(* IEC 61131-3 sources: plc-process-lib/src/POUs/Devices/FB_Valve, 28 files *)

(* ---- FB_Valve.decl.st ---- *)
// Назначение: запорная арматура двух видов. Задвижка с электроприводом (Motorized): выходы
//             «открывать» и «закрывать», стоп в промежутке, смена направления в ходе — через паузу
//             tReverse. Клапан с соленоидом (SolenoidEto, SolenoidEtc): одна катушка, пружинный
//             возврат. Открыть, закрыть, стоп от HMI и от автоматики; концевики ZSO/ZSC (или
//             положение по времени хода), контроль времени хода, «оба концевика», уход с концевика,
//             муфта ограничения момента, внешняя авария; Reset с окном tResetWindow; блокировки с
//             положением безопасности и первопричиной, разрешения по направлениям; режимы Auto,
//             Manual, Local, OutOfService; циклы и время работы привода в stRetain. Блокировка при одних
//             отказах контроля ведёт задвижку в положение безопасности (VLV-20); муфта открытия при
//             страгивании с седла — не заклинивание (VLV-21). Наследует FB_DeviceBase: тело — нормативный
//             порядок цикла (раздел 9.4 контракта).
// Автор:      kr0nsch
// Версия:     0.1.0
// Документ:   docs/fb/FB_Valve.md
FUNCTION_BLOCK FB_Valve EXTENDS FB_DeviceBase
VAR_INPUT
    xAutoOpen    : BOOL;             // запрос автоматики: TRUE — открыть, FALSE — закрыть
    xZso         : BOOL;             // концевик «открыто»
    xZsc         : BOOL;             // концевик «закрыто»
    xTorqueOpen  : BOOL;             // муфта (моментный выключатель) в сторону открытия
    xTorqueClose : BOOL;             // муфта в сторону закрытия
    xExtFault    : BOOL;             // авария привода: тепловое реле, обрыв фазы, авария интегрированного привода
    xLocal       : BOOL;             // «Местное» на приводе или шкафу
    xPowerOk     : BOOL := TRUE;     // напряжение питания привода
    wInterlock   : WORD := 16#0000;  // блокировки: бит = 1 — вести в eSafePos
    wPermitOpen  : WORD := 16#FFFF;  // разрешения на открытие: бит = 1 — разрешено
    wPermitClose : WORD := 16#FFFF;  // разрешения на закрытие: бит = 1 — разрешено
END_VAR
VAR_IN_OUT
    stCmd    : ST_ValveCmd;          // команды HMI/SCADA (GVL_Hmi.st<TAG>Cmd)
    stRetain : ST_DeviceRetain;      // режим, OOS, циклы, время работы привода (GVL_Persist.st<TAG>Retain)
END_VAR
VAR_IN_OUT CONSTANT
    stCfg : ST_ValveCfg;             // параметры (GVL_Persist.st<TAG>Cfg)
END_VAR
VAR_OUTPUT
    xQOpen  : BOOL;                  // Motorized: контактор «открывать»; соленоид — FALSE
    xQClose : BOOL;                  // Motorized: контактор «закрывать»; соленоид — FALSE
    xQCoil  : BOOL;                  // соленоид: катушка; Motorized — FALSE
    xOpened : BOOL;                  // положение «открыто» (по концевику или по времени хода)
    xClosed : BOOL;                  // положение «закрыто»
    stSts   : ST_ValveSts;           // состояние для HMI/SCADA
END_VAR
VAR
    stCfgLkg     : ST_ValveCfg;      // последняя корректная конфигурация (LKG, нормативно)
    // --- состояние и цель ---
    eState       : E_ValveState := E_ValveState.Unknown;        // состояние арматуры
    eTarget      : E_ValveState := E_ValveState.Intermediate;   // цель вызова: Open, Closed; Intermediate — «никуда»
    eManTarget   : E_ValveState := E_ValveState.Intermediate;   // цель Manual: последняя команда оператора
    eSolCmd      : E_ValveState := E_ValveState.Intermediate;  // соленоид: куда держит катушка; Intermediate — нет тока
    eLastEnd     : E_ValveState := E_ValveState.Unknown;        // последнее достигнутое крайнее положение (счёт циклов)
    eLastDir     : E_ValveState := E_ValveState.Intermediate;   // последнее включённое направление привода (выбег)
    xEndByLs     : BOOL;            // положение Open/Closed подтверждено своим концевиком (контроль ухода)
    // --- отказы: фиксируются до Reset (BothLimits — нет) ---
    xFltFailOpen  : BOOL;            // не открылась за tTravel
    xFltFailClose : BOOL;            // не закрылась за tTravel
    xFltPosLost   : BOOL;            // уход с концевика без команды
    xFltTorque    : BOOL;            // муфта в ходе
    xFltExt       : BOOL;            // внешняя авария
    xBothLimits   : BOOL;            // оба концевика дольше tLimitFilter (не фиксируется)
    xResetWin     : BOOL;            // идёт окно Reset: отказы снимаются, как только ушла причина
    // --- блокировки ---
    wIlkPrev      : WORD;            // блокировки после маски в прошлом вызове (первопричина)
    uiFirstOut    : UINT := GVL_Const.NO_FIRST_OUT;   // номер бита первой блокировки; NO_FIRST_OUT — нет
    // --- время работы привода ---
    xActPrev      : BOOL;            // в прошлом вызове был включён выход привода
    ltActAccum    : LTIME;           // накопитель времени работы привода: доля, меньшая 1 с
    // --- задержки (FB_Delay — единственный таймер библиотеки) ---
    fbTravel      : FB_Delay;        // время хода tTravel: от включения выхода (у соленоида — от смены цели)
    fbReverse     : FB_Delay;        // пауза перед реверсом tReverse
    fbRunOff      : FB_Delay;        // выбег привода: TRUE, пока выход включён, и ещё tReverse после снятия
    fbBoth        : FB_Delay;        // фильтр «оба концевика» tLimitFilter
    fbPosLost     : FB_Delay;        // фильтр ухода с концевика tLimitFilter
    fbResetWin    : FB_Delay;        // окно Reset tResetWindow
    // --- аварийный ход в положение безопасности при отказе контроля (VLV-20) ---
    xSafeMove     : BOOL;            // идёт аварийный ход по блокировке при отказе контроля (Motorized)
    xSafeMoveDone : BOOL;            // аварийный ход закончен: новый — после снятия блокировки или всех отказов
    eSafeDir      : E_ValveState := E_ValveState.Intermediate;   // направление аварийного хода: Opening, Closing
    fbSafeMove    : FB_Delay;        // время аварийного хода tTravel
    // --- страгивание с седла (VLV-21) ---
    xUnseatArmed  : BOOL;            // открытие началось с закрытого положения: муфта при страгивании не отказ
    fbUnseat      : FB_Delay;        // окно страгивания VLV_UNSEAT_BYPASS от начала открытия
    fbZscOff      : FB_Delay;        // ZSC замкнут или разомкнулся меньше tLimitFilter назад
    // --- сигналы и условия этого вызова: считает тело и шаги, читают следующие шаги ---
    xMotorized     : BOOL;           // электропривод (по LKG)
    xAtOpen        : BOOL;           // ZSO подключён и сработал
    xAtClose       : BOOL;           // ZSC подключён и сработал
    xTrqOpen       : BOOL;           // муфта открытия сработала (подключена, Motorized)
    xTrqClose      : BOOL;           // муфта закрытия сработала
    xRemote        : BOOL;           // режим Auto или Manual
    xSupervise     : BOOL;           // контроль концевиков: Auto/Manual и есть корректная Cfg
    xPosSup        : BOOL;           // контроль ухода с концевика: xSupervise и есть напряжение
    wIlk           : WORD;           // блокировки после маски
    xIlkAct        : BOOL;           // блокировка действует (Auto/Manual)
    wPermMissOpen  : WORD;           // недостающие разрешения на открытие
    wPermMissClose : WORD;           // недостающие разрешения на закрытие
    xMayOpen       : BOOL;           // открывать можно: разрешения есть или движение по блокировке
    xMayClose      : BOOL;           // закрывать можно
    xFaultAny      : BOOL;           // есть отказ (фиксированный или «оба концевика»)
    xDrive         : BOOL;           // ПЛК управляет выходами в этом вызове
    xEnterMove     : BOOL;           // в этом вызове началось движение (отсчёт tTravel заново)
END_VAR
VAR_TEMP
    eRes        : E_CmdResult;       // результат ProcessMode
    wPermMiss   : WORD;              // недостающие разрешения для текущего направления
    lrRemain_s  : LREAL;             // остаток времени хода, с
    udiRemain_s : UDINT;             // то же, целые секунды вверх
    xMaint      : BOOL;              // достигнут интервал ТО по циклам
    xAvailDev   : BOOL;              // готовность для автоматики (без учёта Cfg)
    wFltBits    : WORD;              // wFault
    wWrnBits    : WORD;              // wWarning
    wLowBits    : WORD;              // младший байт wStatus
    eDevSt      : E_Ne107Status;     // вклад устройства в NE 107
END_VAR

(* ---- CheckConfig.method.decl.st ---- *)
// Проверка конфигурации: биты wCfgErr арматуры (VLV_CFG_*). Только считает, ничего не меняет
METHOD PROTECTED CheckConfig : WORD
VAR_IN_OUT CONSTANT
    stCfgIn : ST_ValveCfg;   // проверяемая конфигурация
END_VAR
VAR
    wErr      : WORD;        // непройденные проверки
    xMotor    : BOOL;        // электропривод
    xSolenoid : BOOL;        // соленоид любого вида
END_VAR

(* ---- CheckConfig.method.impl.st ---- *)
xMotor := stCfgIn.eType = E_ValveType.Motorized;
xSolenoid := stCfgIn.eType = E_ValveType.SolenoidEto OR stCfgIn.eType = E_ValveType.SolenoidEtc;
IF NOT xMotor AND NOT xSolenoid THEN
    wErr := wErr OR GVL_Const.VLV_CFG_TYPE;
END_IF
IF stCfgIn.tTravel <= T#0S THEN
    wErr := wErr OR GVL_Const.VLV_CFG_TRAVEL;
END_IF
IF (stCfgIn.eSafePos <> E_ValveSafePos.Closed AND stCfgIn.eSafePos <> E_ValveSafePos.Open
    AND stCfgIn.eSafePos <> E_ValveSafePos.Stay)
   OR (xSolenoid AND stCfgIn.eSafePos = E_ValveSafePos.Stay)
THEN
    wErr := wErr OR GVL_Const.VLV_CFG_SAFE_POS;
END_IF
IF (stCfgIn.xCloseOnTorque AND NOT stCfgIn.xTorqueUsed) OR (xSolenoid AND stCfgIn.xTorqueUsed) THEN
    wErr := wErr OR GVL_Const.VLV_CFG_TORQUE;
END_IF
IF xMotor AND stCfgIn.tReverse <= T#0S THEN
    wErr := wErr OR GVL_Const.VLV_CFG_REVERSE;
END_IF
IF stCfgIn.tResetWindow <= T#0S THEN
    wErr := wErr OR GVL_Const.VLV_CFG_RESET;
END_IF
IF NOT CheckAlarmCfg(astCfg := stCfgIn.astAlarm) THEN
    wErr := wErr OR GVL_Const.VLV_CFG_ALARM;
END_IF
CheckConfig := wErr;

(* ---- CountOperations.method.decl.st ---- *)
// Шаг 6.9: циклы «открыто» и время работы привода в stRetain (параметр VAR_IN_OUT, R2).
// Шаг тела FB_Valve; внутренний: PROTECTED (правило L5 контракта), имя зарезервировано для наследников
METHOD PROTECTED CountOperations
VAR_IN_OUT
    stValveRet : ST_DeviceRetain;   // stRetain устройства
END_VAR

(* ---- CountOperations.method.impl.st ---- *)
// 6.9 Счётчики: цикл — вход в Open, если прошлое крайнее положение не Open; время работы — пока
//     включён выход привода (шаг не больше DT_ACCUM_MAX), целые секунды — в stRetain
IF eState = E_ValveState.Open AND eLastEnd <> E_ValveState.Open THEN
    stValveRet.udiOpCount := stValveRet.udiOpCount + 1;
    stValveRet.udiOpCountMaint := stValveRet.udiOpCountMaint + 1;
END_IF
IF eState = E_ValveState.Open OR eState = E_ValveState.Closed THEN
    eLastEnd := eState;
END_IF
IF xActPrev THEN
    ltActAccum := ltActAccum + MIN(ltDt, GVL_Const.DT_ACCUM_MAX);
END_IF
WHILE ltActAccum >= LTIME#1S DO
    ltActAccum := ltActAccum - LTIME#1S;
    stValveRet.udiOpTime_s := stValveRet.udiOpTime_s + 1;
    stValveRet.udiOpTimeMaint_s := stValveRet.udiOpTimeMaint_s + 1;
END_WHILE
xActPrev := xQOpen OR xQClose;

(* ---- CurrentTarget.method.impl.st ---- *)
IF eState = E_ValveState.Opening OR eState = E_ValveState.Open THEN
    CurrentTarget := E_ValveState.Open;
ELSIF eState = E_ValveState.Closing OR eState = E_ValveState.Closed THEN
    CurrentTarget := E_ValveState.Closed;
ELSIF eState = E_ValveState.Reversing THEN
    CurrentTarget := eTarget;
ELSE
    CurrentTarget := E_ValveState.Intermediate;
END_IF

(* ---- DriveToTarget.method.decl.st ---- *)
// Шаг 6.7: переходы движения к цели. Motorized: смена направления в ходе — через Reversing, стоп —
// Intermediate, встречное включение после остановки — не раньше tReverse (выбег); соленоид: смена цели —
// сразу другое направление; муфта в ходе — TorqueTrip, кроме страгивания с седла (VLV-21).
// Шаг тела FB_Valve; внутренний: PROTECTED (правило L5 контракта), имя зарезервировано для наследников
METHOD PROTECTED DriveToTarget
VAR
    xHoldOpen  : BOOL;   // открывать пока нельзя: «закрывать» снят меньше tReverse назад
    xHoldClose : BOOL;   // закрывать пока нельзя: «открывать» снят меньше tReverse назад
    xUnseating : BOOL;   // клин выходит из седла: муфта открытия — не заклинивание (VLV-21)
END_VAR

(* ---- DriveToTarget.method.impl.st ---- *)
// 6.7 Движение к цели. Motorized: смена направления в ходе — через Reversing; стоп — Intermediate.
//     Соленоид: смена цели в ходе — сразу другое направление, стопа нет
xMayOpen := xIlkAct OR wPermMissOpen = 0;
xMayClose := xIlkAct OR wPermMissClose = 0;
xEnterMove := FALSE;
//     выбег: встречное направление включается не раньше tReverse после снятия выхода — и после
//     остановки на концевике или по стопу, а не только при смене направления в ходе. Выходы здесь —
//     прошлого вызова; SetOutputs обновляет fbRunOff выходами этого вызова, поэтому отсчёт идёт ровно
//     от снятия выхода
fbRunOff(xIn := xQOpen OR xQClose, tOffDelay := stCfgLkg.tReverse, itfTime := itfTimeAct);
xHoldOpen := xMotorized AND fbRunOff.xOut AND eLastDir = E_ValveState.Closing;
xHoldClose := xMotorized AND fbRunOff.xOut AND eLastDir = E_ValveState.Opening;
//     страгивание с седла (VLV-21): усилие вырыва клина из седла больше усилия хода, муфта открытия срабатывает при
//     ещё замкнутом ZSC — это не заклинивание (в приводах — шунтирование моментного выключателя при страгивании).
//     Муфта открытия не контролируется, пока ZSC замкнут и ещё tLimitFilter после его размыкания (без ZSC — всё
//     окно), но не дольше VLV_UNSEAT_BYPASS от начала открытия с закрытого положения: клин, который не вышел из
//     седла, даёт TorqueTrip. Контроль заклинивания в ходе остаётся
IF eState <> E_ValveState.Opening THEN
    xUnseatArmed := FALSE;
END_IF
fbZscOff(xIn := xAtClose, tOffDelay := stCfgLkg.tLimitFilter, itfTime := itfTimeAct);
fbUnseat(xIn := xUnseatArmed AND eState = E_ValveState.Opening, tOnDelay := GVL_Const.VLV_UNSEAT_BYPASS,
         itfTime := itfTimeAct);
xUnseating := xUnseatArmed AND eState = E_ValveState.Opening AND NOT fbUnseat.xOut
              AND (fbZscOff.xOut OR NOT stCfgLkg.xZscUsed);
IF xDrive THEN
    IF eState = E_ValveState.Opening THEN
        IF xAtOpen THEN
            eState := E_ValveState.Open;
        ELSIF xTrqOpen AND NOT xUnseating THEN
            xFltTorque := TRUE;                // момент раньше концевика: заклинивание
            eState := E_ValveState.Fault;
        ELSIF eTarget = E_ValveState.Closed THEN
            IF xMotorized THEN
                eState := E_ValveState.Reversing;
            ELSIF xMayClose THEN
                eState := E_ValveState.Closing;
                xEnterMove := TRUE;
            END_IF
        ELSIF eTarget = E_ValveState.Intermediate AND xMotorized THEN
            eState := E_ValveState.Intermediate;
        END_IF
    ELSIF eState = E_ValveState.Closing THEN
        IF (xAtClose AND NOT stCfgLkg.xCloseOnTorque)
           OR (stCfgLkg.xCloseOnTorque AND xTrqClose AND (xAtClose OR NOT stCfgLkg.xZscUsed))
        THEN
            // по ZSC; при закрытии «по моменту» (клиновая задвижка) — только по муфте: ZSC стоит чуть
            // раньше посадки клина и выход не снимает, иначе задвижка не дожата. Муфта раньше
            // подключённого ZSC — не посадка, а заклинивание: TorqueTrip ниже
            eState := E_ValveState.Closed;
        ELSIF xTrqClose THEN
            xFltTorque := TRUE;
            eState := E_ValveState.Fault;
        ELSIF eTarget = E_ValveState.Open THEN
            IF xMotorized THEN
                eState := E_ValveState.Reversing;
            ELSIF xMayOpen THEN
                eState := E_ValveState.Opening;
                xEnterMove := TRUE;
            END_IF
        ELSIF eTarget = E_ValveState.Intermediate AND xMotorized THEN
            eState := E_ValveState.Intermediate;
        END_IF
    ELSIF eState = E_ValveState.Reversing THEN
        IF eTarget = E_ValveState.Intermediate THEN
            eState := E_ValveState.Intermediate;
        END_IF
    ELSIF eTarget = E_ValveState.Open AND eState <> E_ValveState.Open AND xMayOpen AND NOT xHoldOpen THEN
        // открытие с закрытого положения — окно страгивания от этого вызова
        xUnseatArmed := eState = E_ValveState.Closed;
        IF xUnseatArmed THEN
            fbUnseat.Preset(xValue := FALSE);
            fbUnseat(xIn := TRUE, tOnDelay := GVL_Const.VLV_UNSEAT_BYPASS, itfTime := itfTimeAct);
        END_IF
        eState := E_ValveState.Opening;
        xEnterMove := TRUE;
    ELSIF eTarget = E_ValveState.Closed AND eState <> E_ValveState.Closed AND xMayClose AND NOT xHoldClose THEN
        eState := E_ValveState.Closing;
        xEnterMove := TRUE;
    END_IF
END_IF

(* ---- FB_Valve.impl.st ---- *)
// 0. Первый вызов: число слотов тревог и тип устройства (до ProcessMode)
IF xFirstCall THEN
    uiAlarmCount := GVL_Const.VLV_ALARM_COUNT;
    eDevType := E_DeviceType.Valve;
END_IF

// 1. Время
BeginCycle();

// 2. Конфигурация (LKG)
IF AcceptCfg(wErr := CheckConfig(stCfgIn := stCfg)) THEN
    stCfgLkg := stCfg;
END_IF
// сигналы по LKG: концевик учитывается, только если подключён; муфта — только у Motorized
xMotorized := stCfgLkg.eType = E_ValveType.Motorized;
xAtOpen := stCfgLkg.xZsoUsed AND xZso;
xAtClose := stCfgLkg.xZscUsed AND xZsc;
xTrqOpen := xMotorized AND stCfgLkg.xTorqueUsed AND xTorqueOpen;
xTrqClose := xMotorized AND stCfgLkg.xTorqueUsed AND xTorqueClose;

// 3. Reset (метод ResetFaults; бит xReset сбрасывает RunAlarms в шаге 7)
ResetFaults(xRequest := xResetReq OR stCmd.stCommon.xReset);

// 4. Режим: вывод из работы — только когда арматура не движется
eRes := ProcessMode(xLocalSel := xLocal, xLocalSupported := TRUE,
                    xOosAllowed := eState <> E_ValveState.Opening AND eState <> E_ValveState.Closing
                                   AND eState <> E_ValveState.Reversing AND NOT xSafeMove,
                    stCmd := stCmd.stCommon, stRetain := stRetain);
IF eRes <> E_CmdResult.None THEN
    SetCmdResult(eResult := eRes);
END_IF

// 5. Условия вызова для шагов-методов; команды устройства (метод HandleCommands)
xRemote := eMode = E_DeviceMode.Auto OR eMode = E_DeviceMode.Manual;
wIlk := wInterlock AND stCfgLkg.wInterlockMask;
xIlkAct := xRemote AND wIlk <> 0;
wPermMissOpen := stCfgLkg.wPermitOpenMask AND NOT wPermitOpen;
wPermMissClose := stCfgLkg.wPermitCloseMask AND NOT wPermitClose;
xFaultAny := xFltFailOpen OR xFltFailClose OR xFltPosLost OR xFltTorque OR xFltExt OR xBothLimits;
HandleCommands(stValveCmd := stCmd, stValveRet := stRetain);

// 6. Логика по stCfgLkg: цель, контроль концевиков, состояние, движение, выходы, счётчики
SelectTarget();
SuperviseLimits();
TrackPosition();
DriveToTarget();
RunTravelTimers();
SafeMoveOnFault();
SetOutputs();
CountOperations(stValveRet := stRetain);

// 7. Тревоги (слоты E_ValveAlarm)
axAlmCond[E_ValveAlarm.FailToOpen] := xFltFailOpen;
axAlmCond[E_ValveAlarm.FailToClose] := xFltFailClose;
axAlmCond[E_ValveAlarm.BothLimits] := xBothLimits;
axAlmCond[E_ValveAlarm.PositionLost] := xFltPosLost;
axAlmCond[E_ValveAlarm.TorqueTrip] := xFltTorque;
axAlmCond[E_ValveAlarm.ExtFault] := xFltExt;
axAlmCond[E_ValveAlarm.InterlockAct] := xIlkAct;
RunAlarms(udiIdBase := stCfgLkg.udiAlarmIdBase, stCmd := stCmd.stCommon, astCfg := stCfgLkg.astAlarm);

// 8. Состояние
IF xRemote AND NOT xIlkAct AND eTarget = E_ValveState.Open AND eState <> E_ValveState.Open THEN
    wPermMiss := wPermMissOpen;
ELSIF xRemote AND NOT xIlkAct AND eTarget = E_ValveState.Closed AND eState <> E_ValveState.Closed THEN
    wPermMiss := wPermMissClose;
ELSE
    wPermMiss := 0;
END_IF
IF eState = E_ValveState.Opening OR eState = E_ValveState.Closing OR xSafeMove THEN
    // остаток до таймаута хода (аварийного хода), целые секунды вверх, не больше UINT_MAX
    IF xSafeMove THEN
        lrRemain_s := F_TimeToSec(tIn := fbSafeMove.tRemaining);
    ELSE
        lrRemain_s := F_TimeToSec(tIn := fbTravel.tRemaining);
    END_IF
    udiRemain_s := LREAL_TO_UDINT(lrRemain_s);
    IF UDINT_TO_LREAL(udiRemain_s) < lrRemain_s THEN
        udiRemain_s := udiRemain_s + 1;
    END_IF
    stSts.uiTravelRemain_s := UDINT_TO_UINT(MIN(udiRemain_s, UINT_TO_UDINT(GVL_Const.UINT_MAX)));
ELSE
    stSts.uiTravelRemain_s := 0;
END_IF
xMaint := stCfgLkg.udiMaintCycles > 0 AND stRetain.udiOpCountMaint >= stCfgLkg.udiMaintCycles;
wFltBits := SEL(xFltFailOpen, 0, GVL_Const.VLV_FLT_FAIL_TO_OPEN)
            OR SEL(xFltFailClose, 0, GVL_Const.VLV_FLT_FAIL_TO_CLOSE)
            OR SEL(xBothLimits, 0, GVL_Const.VLV_FLT_BOTH_LIMITS)
            OR SEL(xFltPosLost, 0, GVL_Const.VLV_FLT_POSITION_LOST)
            OR SEL(xFltTorque, 0, GVL_Const.VLV_FLT_TORQUE_TRIP)
            OR SEL(xFltExt, 0, GVL_Const.VLV_FLT_EXT_FAULT);
wWrnBits := SEL(xMaint, 0, GVL_Const.VLV_WRN_MAINT_CYCLES)
            OR SEL(xPowerOk, GVL_Const.VLV_WRN_POWER_LOST, 0)
            OR SEL(eMode = E_DeviceMode.Local AND wIlk <> 0, 0, GVL_Const.VLV_WRN_INTERLOCK_IN_LOCAL)
            OR SEL((eState = E_ValveState.Open AND NOT stCfgLkg.xZsoUsed)
                   OR (eState = E_ValveState.Closed AND NOT stCfgLkg.xZscUsed AND NOT stCfgLkg.xCloseOnTorque),
                   0, GVL_Const.VLV_WRN_POSITION_BY_TIME)
            OR SEL(eState = E_ValveState.Unknown, 0, GVL_Const.VLV_WRN_POSITION_UNKNOWN);
xAvailDev := eMode = E_DeviceMode.Auto AND wFltBits = 0 AND wIlk = 0 AND xPowerOk;
wLowBits := SEL(xOpened, 0, GVL_Const.VLV_STS_OPENED)
            OR SEL(xClosed, 0, GVL_Const.VLV_STS_CLOSED)
            OR SEL(eState = E_ValveState.Opening OR (xSafeMove AND eSafeDir = E_ValveState.Opening), 0,
                   GVL_Const.VLV_STS_OPENING)
            OR SEL(eState = E_ValveState.Closing OR (xSafeMove AND eSafeDir = E_ValveState.Closing), 0,
                   GVL_Const.VLV_STS_CLOSING)
            OR SEL(xIlkAct, 0, GVL_Const.VLV_STS_INTERLOCKED)
            OR SEL(wPermMiss <> 0, 0, GVL_Const.VLV_STS_PERMIT_MISSING)
            OR SEL(xTrqOpen OR xTrqClose, 0, GVL_Const.VLV_STS_TORQUE)
            OR SEL(xAvailDev AND xCfgEverOk, 0, GVL_Const.VLV_STS_AVAILABLE);
IF wFltBits <> 0 THEN
    eDevSt := E_Ne107Status.Failure;
ELSIF xMaint THEN
    eDevSt := E_Ne107Status.MaintenanceRequired;
ELSE
    eDevSt := E_Ne107Status.Good;
END_IF
stSts.eState := eState;
stSts.wInterlock := wIlk;
stSts.wPermitMissing := wPermMiss;
stSts.uiFirstOut := uiFirstOut;
stSts.wReserve := 0;
stSts.udiCycles := stRetain.udiOpCount;
stSts.udiCyclesMaint := stRetain.udiOpCountMaint;
stSts.rActTime_h := LREAL_TO_REAL(UDINT_TO_LREAL(stRetain.udiOpTime_s) / UDINT_TO_LREAL(GVL_Const.S_PER_H));
FinishCycle(eDevStatus := eDevSt, xAvailableDev := xAvailDev, wLow := wLowBits, wFaultBits := wFltBits,
            wWarnBits := wWrnBits, stCommon := stSts.stCommon);

(* ---- HandleCommands.method.decl.st ---- *)
// Шаг 5: команды HMI xClose > xOpen > xStop и xResetMaint; результат каждой — SetCmdResult. В Auto
// принятая команда переводит в Manual (оператор вмешался — автомат отпущен). Структуры — параметрами
// VAR_IN_OUT: метод не обращается к VAR_IN_OUT экземпляра (R2).
// Шаг тела FB_Valve; внутренний: PROTECTED (правило L5 контракта), имя зарезервировано для наследников
METHOD PROTECTED HandleCommands
VAR_IN_OUT
    stValveCmd : ST_ValveCmd;       // stCmd устройства: импульсы сбрасываются
    stValveRet : ST_DeviceRetain;   // stRetain устройства: режим, счётчики «с ТО»
END_VAR
VAR
    eCmdTgt : E_ValveState := E_ValveState.Intermediate;   // цель команды; Intermediate — стоп
    eResCmd : E_CmdResult := E_CmdResult.None;             // результат команды
END_VAR

(* ---- HandleCommands.method.impl.st ---- *)
IF stValveCmd.xClose OR stValveCmd.xOpen OR stValveCmd.xStop THEN
    IF stValveCmd.xClose THEN
        eCmdTgt := E_ValveState.Closed;
    ELSIF stValveCmd.xOpen THEN
        eCmdTgt := E_ValveState.Open;
    ELSE
        eCmdTgt := E_ValveState.Intermediate;
    END_IF
    IF NOT xRemote THEN
        eResCmd := E_CmdResult.RejectedMode;
    ELSIF eCmdTgt = E_ValveState.Intermediate THEN
        // стоп: только у электропривода; безопасен, поэтому без проверки Cfg и отказов
        IF NOT xMotorized THEN
            eResCmd := E_CmdResult.RejectedNotSupported;
        ELSIF xIlkAct THEN
            eResCmd := E_CmdResult.RejectedInterlock;
        ELSE
            eResCmd := E_CmdResult.Accepted;
        END_IF
    ELSIF NOT xCfgEverOk THEN
        eResCmd := E_CmdResult.RejectedCfg;
    ELSIF xFaultAny THEN
        eResCmd := E_CmdResult.RejectedFault;
    ELSIF xIlkAct THEN
        eResCmd := E_CmdResult.RejectedInterlock;
    ELSIF (eCmdTgt = E_ValveState.Open AND wPermMissOpen <> 0)
          OR (eCmdTgt = E_ValveState.Closed AND wPermMissClose <> 0)
    THEN
        eResCmd := E_CmdResult.RejectedPermit;
    ELSIF NOT xPowerOk THEN
        eResCmd := E_CmdResult.RejectedInhibit;
    ELSE
        eResCmd := E_CmdResult.Accepted;
    END_IF
    IF eResCmd = E_CmdResult.Accepted THEN
        // Auto -> Manual (хук: цель := текущее направление); в Manual режим не меняется
        SwitchRemoteMode(eNew := E_DeviceMode.Manual, stRetain := stValveRet);
        eManTarget := eCmdTgt;
    END_IF
    SetCmdResult(eResult := eResCmd);
END_IF
stValveCmd.xOpen := FALSE;
stValveCmd.xClose := FALSE;
stValveCmd.xStop := FALSE;
IF stValveCmd.xResetMaint THEN
    stValveRet.udiOpCountMaint := 0;
    stValveRet.udiOpTimeMaint_s := 0;
    SetCmdResult(eResult := E_CmdResult.Accepted);
    stValveCmd.xResetMaint := FALSE;
END_IF

(* ---- LimitPosition.method.decl.st ---- *)
// Положение по концевикам (с учётом «подключён»): только ZSO — Open, только ZSC — Closed, оба —
// Unknown; ни одного — Intermediate, а без концевиков — Unknown. Старт ПЛК и снятие отказа.
// Внутренний шаг устройства: PROTECTED (правило L5 контракта), имя зарезервировано для наследников
METHOD PROTECTED LimitPosition : E_ValveState
VAR
    xOpenLs  : BOOL;   // ZSO подключён и сработал
    xCloseLs : BOOL;   // ZSC подключён и сработал
END_VAR

(* ---- LimitPosition.method.impl.st ---- *)
xOpenLs := stCfgLkg.xZsoUsed AND xZso;
xCloseLs := stCfgLkg.xZscUsed AND xZsc;
IF xOpenLs AND xCloseLs THEN
    LimitPosition := E_ValveState.Unknown;
ELSIF xOpenLs THEN
    LimitPosition := E_ValveState.Open;
ELSIF xCloseLs THEN
    LimitPosition := E_ValveState.Closed;
ELSIF stCfgLkg.xZsoUsed OR stCfgLkg.xZscUsed THEN
    LimitPosition := E_ValveState.Intermediate;
ELSE
    LimitPosition := E_ValveState.Unknown;
END_IF

(* ---- OnModeChanged.method.decl.st ---- *)
// Хук смены режима: сначала база (SUPER^); переход в Manual — цель := текущее направление или
// положение (арматура не дёргается); вход в OutOfService снимает зафиксированные отказы и
// первопричину. VAR_IN_OUT устройства не трогает (R2)
METHOD PROTECTED OnModeChanged
VAR_INPUT
    eOld : E_DeviceMode;   // режим до смены
    eNew : E_DeviceMode;   // новый режим
END_VAR

(* ---- OnModeChanged.method.impl.st ---- *)
SUPER^.OnModeChanged(eOld := eOld, eNew := eNew);
IF eNew = E_DeviceMode.Manual THEN
    eManTarget := CurrentTarget();
END_IF
IF eNew = E_DeviceMode.OutOfService THEN
    xFltFailOpen := FALSE;
    xFltFailClose := FALSE;
    xFltPosLost := FALSE;
    xFltTorque := FALSE;
    xFltExt := FALSE;
    xResetWin := FALSE;
    uiFirstOut := GVL_Const.NO_FIRST_OUT;
END_IF

(* ---- ResetFaults.method.decl.st ---- *)
// Шаг 3: Reset. Результат Accepted сразу; в окне tResetWindow зафиксированные отказы снимаются, как
// только ушла их причина (ход и положение — сразу: привод стоит); если к концу окна отказ остался —
// второй результат RejectedFault. Первопричина блокировки снимается.
// Шаг тела FB_Valve; внутренний: PROTECTED (правило L5 контракта), имя зарезервировано для наследников
METHOD PROTECTED ResetFaults
VAR_INPUT
    xRequest : BOOL;   // Reset() или stCmd.stCommon.xReset в этом вызове
END_VAR

(* ---- ResetFaults.method.impl.st ---- *)
IF xRequest THEN
    uiFirstOut := GVL_Const.NO_FIRST_OUT;
    SetCmdResult(eResult := E_CmdResult.Accepted);
    IF xFltFailOpen OR xFltFailClose OR xFltPosLost OR xFltTorque OR xFltExt THEN
        xResetWin := TRUE;
        fbResetWin.Preset(xValue := FALSE);
    END_IF
END_IF
fbResetWin(xIn := xResetWin, tOnDelay := stCfgLkg.tResetWindow, itfTime := itfTimeAct);
IF xResetWin THEN
    // отказы хода и положения: привод стоит, причина в прошлом — снимаются сразу
    xFltFailOpen := FALSE;
    xFltFailClose := FALSE;
    xFltPosLost := FALSE;
    IF NOT xTrqOpen AND NOT xTrqClose THEN
        xFltTorque := FALSE;
    END_IF
    IF NOT xExtFault THEN
        xFltExt := FALSE;
    END_IF
    IF NOT xFltTorque AND NOT xFltExt THEN
        xResetWin := FALSE;
    ELSIF fbResetWin.xOut THEN
        SetCmdResult(eResult := E_CmdResult.RejectedFault);
        xResetWin := FALSE;
    END_IF
END_IF

(* ---- RunTravelTimers.method.impl.st ---- *)
//     пауза реверса: отсчёт с входа в Reversing, затем направление по цели
fbReverse(xIn := eState = E_ValveState.Reversing, tOnDelay := stCfgLkg.tReverse, itfTime := itfTimeAct);
IF eState = E_ValveState.Reversing AND fbReverse.xOut THEN
    IF eTarget = E_ValveState.Open AND xMayOpen THEN
        eState := E_ValveState.Opening;
        xEnterMove := TRUE;
    ELSIF eTarget = E_ValveState.Closed AND xMayClose THEN
        eState := E_ValveState.Closing;
        xEnterMove := TRUE;
    ELSE
        eState := E_ValveState.Intermediate;
    END_IF
END_IF
//     время хода: отсчёт заново с каждого начала движения. Концевик положения подключён (у
//     закрытия — или закрытие по моменту) — таймаут = отказ; не подключён — положение по времени
IF xEnterMove THEN
    fbTravel.Preset(xValue := FALSE);
END_IF
fbTravel(xIn := eState = E_ValveState.Opening OR eState = E_ValveState.Closing, tOnDelay := stCfgLkg.tTravel,
         itfTime := itfTimeAct);
IF fbTravel.xOut THEN
    IF eState = E_ValveState.Opening THEN
        IF stCfgLkg.xZsoUsed THEN
            xFltFailOpen := TRUE;
            eState := E_ValveState.Fault;
        ELSE
            eState := E_ValveState.Open;
        END_IF
    ELSIF eState = E_ValveState.Closing THEN
        IF stCfgLkg.xZscUsed OR stCfgLkg.xCloseOnTorque THEN
            xFltFailClose := TRUE;
            eState := E_ValveState.Fault;
        ELSE
            eState := E_ValveState.Closed;
        END_IF
    END_IF
END_IF

//     крайнее положение подтверждено концевиком (по времени хода и «по моменту» — нет): только
//     такое положение контролируется на уход с концевика
IF (eState = E_ValveState.Open AND xAtOpen) OR (eState = E_ValveState.Closed AND xAtClose) THEN
    xEndByLs := TRUE;
ELSIF eState <> E_ValveState.Open AND eState <> E_ValveState.Closed THEN
    xEndByLs := FALSE;
END_IF

(* ---- SafeMoveOnFault.method.decl.st ---- *)
// Шаг 6.7а (VLV-20): аварийный ход в положение безопасности по блокировке, когда отказали только средства
// контроля (BothLimits, PositionLost, FailToOpen, FailToClose), а привод исправен: защита важнее диагностики.
// Только Motorized (соленоид при отказе уходит на пружину, A-10), с положением безопасности Open или Closed; не
// при внешней аварии, муфте, без напряжения и без корректной Cfg. Концевикам при отказе контроля верить нельзя:
// ход заканчивается по согласованному концевику положения безопасности (свой замкнут, встречный нет), по муфте в
// этом направлении или через tTravel. Пока блокировка и отказ держатся, ход не повторяется. Начало — после выбега
// встречного направления (VLV-05).
// Шаг тела FB_Valve; внутренний: PROTECTED (правило L5 контракта), имя зарезервировано для наследников
METHOD PROTECTED SafeMoveOnFault
VAR
    xMayMove : BOOL;   // аварийный ход допустим в этом вызове
    xEnd     : BOOL;   // аварийный ход закончен в этом вызове
END_VAR

(* ---- SafeMoveOnFault.method.impl.st ---- *)
xMayMove := xMotorized AND xIlkAct AND xFaultAny AND xCfgEverOk AND xPowerOk AND NOT xFltExt AND NOT xFltTorque
            AND (stCfgLkg.eSafePos = E_ValveSafePos.Open OR stCfgLkg.eSafePos = E_ValveSafePos.Closed);
IF NOT xMayMove THEN
    xSafeMove := FALSE;
    IF NOT (xIlkAct AND xFaultAny) THEN
        // блокировка или отказы сняты: следующий эпизод — новый аварийный ход
        xSafeMoveDone := FALSE;
    END_IF
ELSIF NOT xSafeMove AND NOT xSafeMoveDone THEN
    IF stCfgLkg.eSafePos = E_ValveSafePos.Closed AND NOT (fbRunOff.xOut AND eLastDir = E_ValveState.Opening) THEN
        eSafeDir := E_ValveState.Closing;
        xSafeMove := TRUE;
    ELSIF stCfgLkg.eSafePos = E_ValveSafePos.Open AND NOT (fbRunOff.xOut AND eLastDir = E_ValveState.Closing) THEN
        eSafeDir := E_ValveState.Opening;
        xSafeMove := TRUE;
    END_IF
    IF xSafeMove THEN
        fbSafeMove.Preset(xValue := FALSE);
    END_IF
END_IF
fbSafeMove(xIn := xSafeMove, tOnDelay := stCfgLkg.tTravel, itfTime := itfTimeAct);
IF xSafeMove THEN
    IF eSafeDir = E_ValveState.Closing THEN
        xEnd := (xAtClose AND NOT xAtOpen) OR xTrqClose;
    ELSE
        xEnd := (xAtOpen AND NOT xAtClose) OR xTrqOpen;
    END_IF
    IF xEnd OR fbSafeMove.xOut THEN
        xSafeMove := FALSE;
        xSafeMoveDone := TRUE;
    END_IF
END_IF

(* ---- SelectTarget.method.decl.st ---- *)
// Шаг 6.1–6.2: цель вызова (Auto — запрос автоматики, Manual — команда оператора, Local/OOS — нет,
// блокировка — положение безопасности) и первопричина блокировки.
// Шаг тела FB_Valve; внутренний: PROTECTED (правило L5 контракта), имя зарезервировано для наследников
METHOD PROTECTED SelectTarget
VAR
    wBit  : WORD;   // бит при поиске первопричины
    uiBit : UINT;   // номер бита
END_VAR

(* ---- SelectTarget.method.impl.st ---- *)
// 6.1 Цель: Auto — по запросу автоматики, Manual — по команде оператора, Local/OOS — нет;
//     блокировка (Auto/Manual) — положение безопасности (Stay — стоп)
IF eMode = E_DeviceMode.Auto THEN
    IF xAutoOpen THEN
        eTarget := E_ValveState.Open;
    ELSE
        eTarget := E_ValveState.Closed;
    END_IF
ELSIF eMode = E_DeviceMode.Manual THEN
    eTarget := eManTarget;
ELSE
    eTarget := E_ValveState.Intermediate;
END_IF
IF xIlkAct THEN
    IF stCfgLkg.eSafePos = E_ValveSafePos.Open THEN
        eTarget := E_ValveState.Open;
    ELSIF stCfgLkg.eSafePos = E_ValveSafePos.Closed THEN
        eTarget := E_ValveState.Closed;
    ELSE
        eTarget := E_ValveState.Intermediate;
    END_IF
    // блокировка не фиксируется: после её снятия Manual остаётся в положении безопасности
    IF eMode = E_DeviceMode.Manual THEN
        eManTarget := eTarget;
    END_IF
END_IF

// 6.2 Первопричина: при переходе слова блокировок из 0 в не 0 — номер младшего взведённого бита
//     (держится до Reset или входа в OutOfService). Цикл конечен: wIlk <> 0
IF wIlkPrev = 0 AND wIlk <> 0 AND eMode <> E_DeviceMode.OutOfService THEN
    wBit := 1;
    uiBit := 0;
    WHILE (wIlk AND wBit) = 0 DO
        wBit := SHL(wBit, 1);
        uiBit := uiBit + 1;
    END_WHILE
    uiFirstOut := uiBit;
END_IF
wIlkPrev := wIlk;

(* ---- SetOutputs.method.decl.st ---- *)
// Шаг 6.8: выходы привода и катушки, положение для логики. Без управления и при отказе выходы сняты,
// катушка обесточена (положение пружины); при отказе контроля — аварийный ход по блокировке (VLV-20).
// Шаг тела FB_Valve; внутренний: PROTECTED (правило L5 контракта), имя зарезервировано для наследников
METHOD PROTECTED SetOutputs
VAR
    xOutEn : BOOL;   // выходы разрешены
END_VAR

(* ---- SetOutputs.method.impl.st ---- *)
// 6.8 Выходы. Без управления и при отказе выходы сняты, катушка обесточена (положение пружины)
IF NOT xDrive OR eState = E_ValveState.Fault OR xMotorized THEN
    eSolCmd := E_ValveState.Intermediate;
ELSIF eState = E_ValveState.Opening OR (eState = E_ValveState.Open AND eTarget = E_ValveState.Open) THEN
    eSolCmd := E_ValveState.Open;
ELSIF eState = E_ValveState.Closing OR (eState = E_ValveState.Closed AND eTarget = E_ValveState.Closed) THEN
    eSolCmd := E_ValveState.Closed;
END_IF
xOutEn := xDrive AND eState <> E_ValveState.Fault;
//     аварийный ход в положение безопасности (VLV-20) — только при отказе (eState = Fault): с обычными выходами не
//     пересекается
xQOpen := (xOutEn AND xMotorized AND eState = E_ValveState.Opening)
          OR (xSafeMove AND eSafeDir = E_ValveState.Opening);
xQClose := (xOutEn AND xMotorized AND eState = E_ValveState.Closing)
           OR (xSafeMove AND eSafeDir = E_ValveState.Closing);
xQCoil := xOutEn AND ((stCfgLkg.eType = E_ValveType.SolenoidEto AND eSolCmd = E_ValveState.Open)
                      OR (stCfgLkg.eType = E_ValveType.SolenoidEtc AND eSolCmd = E_ValveState.Closed));
xOpened := eState = E_ValveState.Open OR (eState = E_ValveState.Fault AND xAtOpen AND NOT xAtClose);
xClosed := eState = E_ValveState.Closed OR (eState = E_ValveState.Fault AND xAtClose AND NOT xAtOpen);
//     выбег привода: последнее включённое направление и отсчёт tReverse от снятия выхода (DriveToTarget)
IF xQOpen THEN
    eLastDir := E_ValveState.Opening;
ELSIF xQClose THEN
    eLastDir := E_ValveState.Closing;
END_IF
fbRunOff(xIn := xQOpen OR xQClose, tOffDelay := stCfgLkg.tReverse, itfTime := itfTimeAct);

(* ---- SuperviseLimits.method.decl.st ---- *)
// Шаг 6.3–6.4: внешняя авария, «оба концевика», уход с концевика (фильтры tLimitFilter).
// Шаг тела FB_Valve; внутренний: PROTECTED (правило L5 контракта), имя зарезервировано для наследников
METHOD PROTECTED SuperviseLimits
VAR
    xLeftEnd : BOOL;   // в Open/Closed, подтверждённом концевиком, он пропал
END_VAR

(* ---- SuperviseLimits.method.impl.st ---- *)
// 6.3 Внешняя авария: во всех режимах, кроме OutOfService; фиксируется
IF xExtFault AND eMode <> E_DeviceMode.OutOfService THEN
    xFltExt := TRUE;
END_IF

// 6.4 Концевики (контроль — в Auto/Manual при корректной Cfg; в Local и OOS арматуру двигают руками).
//     «Оба концевика» дольше tLimitFilter — нефиксируемый отказ; при старте ПЛК — сразу
xSupervise := xRemote AND xCfgEverOk;
fbBoth(xIn := xSupervise AND xAtOpen AND xAtClose, tOnDelay := stCfgLkg.tLimitFilter, itfTime := itfTimeAct);
IF xFirstCall THEN
    fbBoth.Preset(xValue := xSupervise AND xAtOpen AND xAtClose);
END_IF
xBothLimits := fbBoth.xOut;
//     уход с концевика: в Open/Closed, подтверждённом концевиком, он пропал без команды дольше
//     tLimitFilter — фиксируемый отказ; без напряжения не контролируется (соленоид уходит на пружину)
xPosSup := xSupervise AND xPowerOk;
xLeftEnd := xEndByLs AND ((eState = E_ValveState.Open AND NOT xAtOpen)
                          OR (eState = E_ValveState.Closed AND NOT xAtClose));
fbPosLost(xIn := xPosSup AND xLeftEnd, tOnDelay := stCfgLkg.tLimitFilter, itfTime := itfTimeAct);
IF fbPosLost.xOut THEN
    xFltPosLost := TRUE;
END_IF

(* ---- TrackPosition.method.decl.st ---- *)
// Шаг 6.5–6.6: отказ и его снятие, старт ПЛК, останов без управления; без движения — состояние по
// концевикам.
// Шаг тела FB_Valve; внутренний: PROTECTED (правило L5 контракта), имя зарезервировано для наследников
METHOD PROTECTED TrackPosition
VAR
    xLeftEnd : BOOL;   // в Open/Closed, подтверждённом концевиком, он пропал
    xCoilEnd : BOOL;   // соленоид в положении, которое держит ток катушки (Eto — Open, Etc — Closed)
END_VAR

(* ---- TrackPosition.method.impl.st ---- *)
// 6.5 Автомат состояний: отказ, снятие отказа, останов без управления
xFaultAny := xFltFailOpen OR xFltFailClose OR xFltPosLost OR xFltTorque OR xFltExt OR xBothLimits;
xDrive := xRemote AND xCfgEverOk AND xPowerOk AND NOT xFaultAny;
IF xFirstCall THEN
    // старт ПЛК: состояние по концевикам; Manual: цель := текущее положение
    eState := LimitPosition();
    IF eState = E_ValveState.Open OR eState = E_ValveState.Closed THEN
        eLastEnd := eState;
    END_IF
    eManTarget := CurrentTarget();
END_IF
IF xFaultAny THEN
    eState := E_ValveState.Fault;
    eManTarget := E_ValveState.Intermediate;   // после Reset арматура в Manual сама не двинется
ELSIF eState = E_ValveState.Fault THEN
    eState := LimitPosition();                 // отказы сняты: далее — по концевикам
ELSIF NOT xDrive AND (eState = E_ValveState.Opening OR eState = E_ValveState.Closing
                      OR eState = E_ValveState.Reversing)
THEN
    eState := E_ValveState.Intermediate;       // выходы сняты: нет напряжения, Local, OOS
END_IF
IF NOT xPowerOk THEN
    eManTarget := E_ValveState.Intermediate;   // нет напряжения: Manual стоит, цель снята
END_IF

// 6.6 Без движения — состояние по концевикам. При контроле уход с концевика и «оба концевика»
//     держат состояние до срабатывания фильтра (дальше — Fault)
IF eState = E_ValveState.Open OR eState = E_ValveState.Closed OR eState = E_ValveState.Intermediate
   OR eState = E_ValveState.Unknown
THEN
    //  положение «по времени» (не подтверждённое своим концевиком) держится, только пока арматурой
    //  управляет ПЛК: в Local и OOS её двигают с места или руками, соленоид без тока катушки уходит на
    //  пружину. Дальше — только по концевикам (без концевиков — Unknown)
    xCoilEnd := (stCfgLkg.eType = E_ValveType.SolenoidEto AND eState = E_ValveState.Open)
                OR (stCfgLkg.eType = E_ValveType.SolenoidEtc AND eState = E_ValveState.Closed);
    IF (eState = E_ValveState.Open OR eState = E_ValveState.Closed) AND NOT xEndByLs
       AND (NOT xRemote OR (xCoilEnd AND NOT xDrive))
    THEN
        eState := LimitPosition();
    END_IF
    xLeftEnd := xEndByLs AND ((eState = E_ValveState.Open AND NOT xAtOpen)
                              OR (eState = E_ValveState.Closed AND NOT xAtClose));
    IF NOT (xLeftEnd AND xPosSup) THEN
        IF xAtOpen AND xAtClose THEN
            IF NOT xSupervise THEN
                eState := E_ValveState.Unknown;
            END_IF
        ELSIF xAtOpen THEN
            eState := E_ValveState.Open;
        ELSIF xAtClose THEN
            eState := E_ValveState.Closed;
        ELSIF xLeftEnd THEN
            eState := E_ValveState.Intermediate;
        END_IF
    END_IF
END_IF
